Fanuc KAREL source: KA00110.KL

PROGRAM KA00110
%NOLOCKGROUP
VAR
  SRC: CONFIG
  DST: REAL
BEGIN
  SRC.CFG_FLIP = TRUE
  DST = SRC
END KA00110
